Staubli VAL3: Algorithm4.pjx

--- Algorithm4.pjx ---
Parameters version=s8.10.5Cs9_BS2172 stackSize=5000 millimeterUnit=true
Program file=_CalpCircle.pgx
Program file=CalAdjustXY2.pgx
Program file=CalAdjustXY3.pgx
Program file=CalToolPos2.pgx
Program file=CalToolPos3.pgx
Program file=CalToolPos6.pgx
Data file=Algorithm4.dtx
Library alias=db path=Disk://SmartTCP_CS9/DataBase4/DataBase4.pjx
Library alias=matrix path=Disk://SmartTCP_CS9/MatrixLib/MatrixLib.pjx

--- Algorithm4.dtx ---
public num nInverseMatrix1[4 4]
  [0,0] = 4.865664
  [0,1] = 0.229739
  [0,2] = 18.957284
  [1,0] = -2.180441
  [1,1] = 5.500387
  [1,2] = 4.336984
  [2,0] = -0.506536
  [2,1] = -1.473409
  [2,2] = -0.0709054
  [3,3] = 1
public num nMatrix1[4 4]
  [0,0] = 0.042143
  [0,1] = -0.196069
  [0,2] = -0.725376
  [1,0] = -0.0165157
  [1,1] = 0.0650218
  [1,2] = -0.43854
  [2,0] = 0.0421337
  [2,1] = 0.0495361
  [2,2] = 0.191493
  [3,3] = 1
public num nMatrix2[4 4]
  [0,0] = 1
  [1,1] = 1
  [2,2] = 1
  [3,0] = 6.816645
  [3,1] = 1120.929616
  [3,2] = 833.829369
  [3,3] = 1
public num nMatrix3[4 4]
  [0,0] = 4.865664
  [0,1] = 0.229739
  [0,2] = 18.957284
  [1,0] = -2.180441
  [1,1] = 5.500387
  [1,2] = 4.336984
  [2,0] = -0.506536
  [2,1] = -1.473409
  [2,2] = -0.0709054
  [3,0] = -2833.317475
  [3,1] = 4938.541162
  [3,2] = 4931.555835
  [3,3] = 1
public num nTeach_3_1[4 4]
  [0,0] = -0.702285
  [0,1] = -0.0819432
  [0,2] = -0.707164
  [1,0] = -0.115862
  [1,1] = 0.993265
  [1,2] = -3.24847E-05
  [2,0] = 0.702404
  [2,1] = 0.0819108
  [2,2] = -0.70705
  [3,0] = 1004.56
  [3,1] = -0.844997
  [3,2] = 227.853426
  [3,3] = 1
public num nTeach_3_2[4 4]
  [0,0] = -0.744428
  [0,1] = 0.279367
  [0,2] = -0.606449
  [1,0] = -0.0993466
  [1,1] = 0.85181
  [1,2] = 0.514345
  [2,0] = 0.66027
  [2,1] = 0.443142
  [2,2] = -0.606357
  [3,0] = 1011.376645
  [3,1] = -59.246821
  [3,2] = 211.566344
  [3,3] = 1
public num nTeach_3_3[4 4]
  [0,0] = -0.879562
  [0,1] = 0.475436
  [0,2] = 0.0182124
  [1,0] = 0.434368
  [1,1] = 0.786788
  [1,2] = 0.438508
  [2,0] = 0.194153
  [2,1] = 0.393606
  [2,2] = -0.898543
  [3,0] = 1061.682795
  [3,1] = -69.818944
  [3,2] = 189.439756
  [3,3] = 1
frame fFrame = {fatherId=world[0]}
num nTeach_2_1[4 4]
num nTeach_2_2[4 4]

--- _CalpCircle.pgx ---
program _CalpCircle(pointRs x_p1, pointRs x_p2, pointRs x_p3, pointRs& x_pCenter, bool& x_bStatus)
  local num x1
  local num y1
  local num x2
  local num y2
  local num x3
  local num y3
  local frame l_fFrame
  local num l_nFrameStatus
  local pointRs l_p3
  local pointRs l_p2
  local pointRs l_p1
  local pointRs l_pCenter
begin
  //圆心算法
  link(l_fFrame,world)
  l_nFrameStatus=setFrame(x_p1,x_p2,x_p3,l_fFrame)
  if l_nFrameStatus!=0
    //3点共线或任意2点过于接近
    popUpMsg("Error!!")
    x_bStatus=false
    return
  endIf
  link(l_p1,l_fFrame)
  link(l_p2,l_fFrame)
  link(l_p3,l_fFrame)
  l_p1.trsf=position(x_p1,l_fFrame)
  l_p2.trsf=position(x_p2,l_fFrame)
  l_p3.trsf=position(x_p3,l_fFrame)
  //
  x1=l_p1.trsf.x
  y1=l_p1.trsf.y
  x2=l_p2.trsf.x
  y2=l_p2.trsf.y
  x3=l_p3.trsf.x
  y3=l_p3.trsf.y
  //
  if((x3-x1)*(y2-y1)-(x2-x1)*(y3-y1))!=0
    link(l_pCenter,l_fFrame)
    l_pCenter.trsf={0,0,0,0,0,0}
    l_pCenter.trsf.x=((y2-y1)*(y3*y3-y1*y1+x3*x3-x1*x1)-(y3-y1)*(y2*y2-y1*y1+x2*x2-x1*x1))/(2*(x3-x1)*(y2-y1)-2*(x2-x1)*(y3-y1))
    l_pCenter.trsf.y=((x2-x1)*(x3*x3-x1*x1+y3*y3-y1*y1)-(x3-x1)*(x2*x2-x1*x1+y2*y2-y1*y1))/(2*(y3-y1)*(x2-x1)-2*(y2-y1)*(x3-x1))
    x_pCenter.trsf=position(l_pCenter,world)
    x_bStatus=true
  else
    x_bStatus=false
    return
 endIf
end

--- CalAdjustXY2.pgx ---
public program CalAdjustXY2()
  local trsf l_trFlange
  local trsf l_trTCP
  local num x
  local num y
  local num z
begin
  //初始化数据
  l_trFlange={0,0,0,0,0,0}
  l_trTCP={0,0,0,0,0,0}
  //计算新的中心位置
  x=(db:pAdjustXY_2_1.trsf.x+db:pAdjustXY_2_2.trsf.x)/2
  y=(db:pAdjustXY_2_1.trsf.y+db:pAdjustXY_2_2.trsf.y)/2
  z=db:pAdjustXY_2_1.trsf.z
  //
  l_trFlange=db:pAdjustXY_2_1.trsf*!db:utCurrentTool.tValue.trsf
  l_trTCP={x,y,z,0,180,0}
  db:tTool2.trsf=!l_trFlange*l_trTCP
  //
  db:tTool2.trsf.rx=db:tTool1.trsf.rx
  db:tTool2.trsf.ry=db:tTool1.trsf.ry
  db:tTool2.trsf.rz=db:tTool1.trsf.rz
  call db:hmiAlert("SaveInTool2","info")
end

--- CalAdjustXY3.pgx ---
public program CalAdjustXY3()
  local trsf l_trFlange
  local trsf l_trTCP
  local num x
  local num y
  local num z
begin
  l_trFlange={0,0,0,0,0,0}
  l_trTCP={0,0,0,0,0,0}
  x=db:pAdjustXY_3_2.trsf.x+db:pAdjustXY_3_3.trsf.x-db:pAdjustXY_3_1.trsf.x
  y=db:pAdjustXY_3_2.trsf.y+db:pAdjustXY_3_3.trsf.y-db:pAdjustXY_3_1.trsf.y
  z=db:pAdjustXY_3_1.trsf.z
  //
  l_trFlange=db:pAdjustXY_3_1.trsf*!db:utCurrentTool.tValue.trsf
  l_trTCP={x,y,z,0,180,0}
  db:tTool2.trsf=!l_trFlange*l_trTCP
  //
  db:tTool2.trsf.rx=db:tTool1.trsf.rx
  db:tTool2.trsf.ry=db:tTool1.trsf.ry
  db:tTool2.trsf.rz=db:tTool1.trsf.rz
  call db:hmiAlert("SaveInTool2","info")
end

--- CalToolPos2.pgx ---
public program CalToolPos2(tool& x_tTool)
  local bool l_bStatus
  local point l_p1
  local num ax1
  local num ax2
  local num ay1
  local num ay2
  local num az1
  local num az2
  local point l_p2
  local trsf l_trP1
  local trsf l_trP2
  local num nx1
  local num nx2
  local num ny1
  local num ny2
  local num nz1
  local num nz2
  local num ox1
  local num ox2
  local num oy1
  local num oy2
  local num oz1
  local num oz2
  local num xf1
  local num xf2
  local num yf1
  local num yf2
  local num zf1
  local num zf2
begin
  //2个带姿态的点求工具值XYZ
  l_trP1=db:pTeach1.trsf
  l_trP2=db:pTeach2.trsf
  //
  //pTeach_2_1转成矩阵nTeach_2_1
  call matrix:Trsf2Matrix(l_trP1,nTeach_2_1)
  //pTeach_2_2转成矩阵nTeach_2_2
  call matrix:Trsf2Matrix(l_trP2,nTeach_2_2)
  //
  //分解矩阵nTeach_2_1
  nx1=nTeach_2_1[0,0]
  ny1=nTeach_2_1[0,1]
  nz1=nTeach_2_1[0,2]
  ox1=nTeach_2_1[1,0]
  oy1=nTeach_2_1[1,1]
  oz1=nTeach_2_1[1,2]
  ax1=nTeach_2_1[2,0]
  ay1=nTeach_2_1[2,1]
  az1=nTeach_2_1[2,2]
  xf1=nTeach_2_1[3,0]
  yf1=nTeach_2_1[3,1]
  zf1=nTeach_2_1[3,2]
  //
  //分解矩阵nTeach_2_2
  nx2=nTeach_2_2[0,0]
  ny2=nTeach_2_2[0,1]
  nz2=nTeach_2_2[0,2]
  ox2=nTeach_2_2[1,0]
  oy2=nTeach_2_2[1,1]
  oz2=nTeach_2_2[1,2]
  ax2=nTeach_2_2[2,0]
  ay2=nTeach_2_2[2,1]
  az2=nTeach_2_2[2,2]
  xf2=nTeach_2_2[3,0]
  yf2=nTeach_2_2[3,1]
  zf2=nTeach_2_2[3,2]
  //
  //***************************************************************************************
  //  │nx1-nx2 , ox1-ox2 ,    0    ,   0  │   │1 , 0 , 0, Tx│   │1 , 0 , 0, xf2-xf1│
  //  │ny2-ny3 , oy2-oy3 ,    0    ,   0  │ * │0 , 1 , 0, Ty│ = │0 , 1 , 0, yf3-yf2│
  //  │nz1-nz3 , oz1-oz3 ,    1    ,   0  │   │0 , 0 , 1, Tz│   │0 , 0 , 1,    0   │
  //  │   0    ,    0    ,    0    ,   1  │   │0 , 0 , 0,  1│   │0 , 0 , 0,    1   │
  //***************************************************************************************
  //构造矩阵nMatrix1
  nMatrix1[0,0]=nx1-nx2
  nMatrix1[0,1]=ny1-ny2
  nMatrix1[0,2]=nz1-nz2
  nMatrix1[0,3]=0
  nMatrix1[1,0]=ox1-ox2
  nMatrix1[1,1]=oy1-oy2
  nMatrix1[1,2]=oz1-oz2
  nMatrix1[1,3]=0
  nMatrix1[2,0]=0
  nMatrix1[2,1]=0
  nMatrix1[2,2]=1
  nMatrix1[2,3]=0
  nMatrix1[3,0]=0
  nMatrix1[3,1]=0
  nMatrix1[3,2]=0
  nMatrix1[3,3]=1
  //
  //构造矩阵nMatrix2
  nMatrix2[0,0]=1
  nMatrix2[0,1]=0
  nMatrix2[0,2]=0
  nMatrix2[0,3]=0

  nMatrix2[1,0]=0
  nMatrix2[1,1]=1
  nMatrix2[1,2]=0
  nMatrix2[1,3]=0

  nMatrix2[2,0]=0
  nMatrix2[2,1]=0
  nMatrix2[2,2]=1
  nMatrix2[2,3]=0

  nMatrix2[3,0]=xf2-xf1
  nMatrix2[3,1]=yf2-yf1
  nMatrix2[3,2]=0
  nMatrix2[3,3]=1
  //***************************************************************************************
  call matrix:InverseMatrix(nMatrix1,nInverseMatrix1,l_bStatus)
  if l_bStatus==false
    //如果nMatrix1不可逆则需重新示教点
    call db:hmiAlert("DeviationIsTooLarge","warning")
  else
    call matrix:MutliMatrix(nInverseMatrix1,nMatrix2,nMatrix3)

    x_tTool.trsf.x=nMatrix3[3,0]
    x_tTool.trsf.y=nMatrix3[3,1]
    x_tTool.trsf.z=0
    x_tTool.trsf.rx=0
    x_tTool.trsf.ry=0
    x_tTool.trsf.rz=0
  endIf
  call db:hmiAlert("SaveInTool1","info")
end

--- CalToolPos3.pgx ---
public program CalToolPos3(tool& x_tTool)
  local bool l_bStatus
  local pointRs l_p1
  local pointRs l_p2
  local pointRs l_p3
  local pointRs l_pCenter
  local tool l_t1
  local tool l_t2
  local tool l_t3
begin
  l_bStatus=false
  link(l_pCenter,world)
  //
  l_p1=db:pTeach1
  l_p2=db:pTeach2
  l_p3=db:pTeach3
  call _CalpCircle(l_p1,l_p2,l_p3,l_pCenter,l_bStatus)
  //

  if l_bStatus==true
    l_pCenter.trsf.rx=0
    l_pCenter.trsf.ry=180
    l_pCenter.trsf.rz=0
  else
    call db:hmiAlert("DeviationIsTooLarge","warning")
  endIf
  l_t1.trsf=!l_p1.trsf*l_pCenter.trsf
  l_t2.trsf=!l_p2.trsf*l_pCenter.trsf
  l_t3.trsf=!l_p3.trsf*l_pCenter.trsf
  x_tTool.trsf.x=(l_t1.trsf.x+l_t2.trsf.x+l_t3.trsf.x)/3
  x_tTool.trsf.y=(l_t1.trsf.y+l_t2.trsf.y+l_t3.trsf.y)/3
  x_tTool.trsf.z=0
  x_tTool.trsf.rx=0
  x_tTool.trsf.ry=0
  x_tTool.trsf.rz=0
  call db:hmiAlert("SaveInTool1","info")
end

--- CalToolPos6.pgx ---
public program CalToolPos6(tool& x_tTool)
  local bool l_bStatus
  local pointRs l_pCenter
  local tool l_t4
  local tool l_t3
  local tool l_t2
  local tool l_t1
  local frame l_fFrame
  local num l_nFrameErr
  local bool l_bBool
  local pointRs l_p5
  local pointRs l_p4
  local pointRs l_p3
  local pointRs l_p2
  local pointRs l_p1
  local pointRs l_p6
begin
  l_bStatus=false
  link(l_pCenter,world)
  //计算中心点坐标
  l_p1=db:pTeach1
  l_p2=db:pTeach2
  l_p3=db:pTeach3
  l_p4=db:pTeach4
  l_p5=db:pTeach5
  l_p6=db:pTeach6
  l_p1.trsf.z=0
  l_p2.trsf.z=0
  l_p3.trsf.z=0
  l_p4.trsf.z=0
  l_p5.trsf.z=0
  l_p6.trsf.z=0
  call _CalpCircle(l_p1,l_p2,l_p3,l_pCenter,l_bStatus)
  //计算工具的xyz
  link(l_p4,world)
  link(l_p5,world)
  link(l_p6,world)
  link(l_fFrame,world)
  l_nFrameErr=setFrame(l_p4,l_p5,l_p6,l_fFrame)
  switch l_nFrameErr
    case 0
      l_pCenter.trsf.rx=l_fFrame.trsf.rx
      l_pCenter.trsf.ry=l_fFrame.trsf.ry
      l_pCenter.trsf.rz=l_fFrame.trsf.rz
      x_tTool.trsf=!l_p4.trsf*l_pCenter.trsf
    break
        case -1,-2
      call db:hmiAlert("DeviationIsTooLarge","info")
    break
  endSwitch
  call db:hmiAlert("SaveInTool1","info")
end
